FUNCTION_BLOCK T_SafeTof_Tests EXTENDS TcUnit.FB_TestSuite
VAR
    // Test_OutputDelayedOff
    group_1 : T_SafeGroup;
    fb_1 : T_SafeTof(group := group_1) := (Parameters := (DelayTime := T#100MS));
    state_1 : INT := 10;
    waitTimer_1 : TON;
    // Test_UnconnectedInputIsRefused
    group_2 : T_SafeGroup;
    fb_2 : T_SafeTof(group := group_2);
END_VAR

Test_OutputDelayedOff();
Test_UnconnectedInputIsRefused();

METHOD PRIVATE Test_OutputDelayedOff
TcUnit.TEST(__POUNAME());
waitTimer_1();

CASE state_1 OF
    10:
        group_1(Run := TRUE);
        fb_1(TofIn1 := TRUE);
        AssertEquals_BOOL(Expected := TRUE, Actual := fb_1.TofOut, Message := 'output on immediately');
        // act
        fb_1(TofIn1 := FALSE);
        AssertEquals_BOOL(Expected := TRUE, Actual := fb_1.TofOut, Message := 'output held during the delay');
        AssertEquals_BYTE(Expected := TO_BYTE(E_SafeFbState.DelayOut), Actual := fb_1.State, Message := 'state DELAYOUT');
        state_1 := 20;
        waitTimer_1(IN := TRUE, PT := T#200MS);
    20:
        group_1(Run := TRUE);
        fb_1(TofIn1 := FALSE);

        IF NOT waitTimer_1.Q THEN
            RETURN;
        END_IF

        waitTimer_1(IN := FALSE);
        // assert
        AssertEquals_BOOL(Expected := FALSE, Actual := fb_1.TofOut, Message := 'output off after the delay');
        TEST_FINISHED_NAMED(__POUNAME());
        state_1 := 10;
END_CASE
END_METHOD

METHOD PRIVATE Test_UnconnectedInputIsRefused
TcUnit.TEST(__POUNAME());
// arrange / act: TofIn1 is unconnected, which the Safety Editor refuses
group_2(Run := TRUE);
fb_2();
group_2(Run := TRUE);
fb_2();
// assert
AssertEquals_BOOL(Expected := TRUE, Actual := fb_2.Error, Message := 'configuration error reported');
AssertEquals_BYTE(Expected := TO_BYTE(E_SafeFbState.Error), Actual := fb_2.State, Message := 'state ERROR');
AssertEquals_WORD(Expected := WORD#16#8000, Actual := fb_2.Diag, Message := 'diag bit 15 configuration refused');
AssertEquals_BOOL(Expected := FALSE, Actual := fb_2.TofOut, Message := 'TofOut stays at its safe value');
AssertEquals_BOOL(Expected := TRUE, Actual := group_2.FbErr, Message := 'the group sees an FB error');
// act: ErrAck 0 -> 1 -> 0 does not clear a configuration error
group_2(Run := TRUE, ErrAck := TRUE);
fb_2();
group_2(Run := TRUE, ErrAck := TRUE);
fb_2();
group_2(Run := TRUE, ErrAck := FALSE);
fb_2();
AssertEquals_BOOL(Expected := TRUE, Actual := fb_2.Error, Message := 'error not acknowledged');
AssertEquals_WORD(Expected := WORD#16#8000, Actual := fb_2.Diag, Message := 'diag bit 15 kept');
TEST_FINISHED_NAMED(__POUNAME());
END_METHOD

END_FUNCTION_BLOCK

(* stored: Version 1.1.0.1
   POU T_SafeTof_Tests: Id {978229da-758b-5bed-80ea-cf07aeecdce2}, SpecialFunc None
   Method Test_OutputDelayedOff: Id {b6d59bd9-12c1-5814-8994-2d4710fe2757}
   Method Test_UnconnectedInputIsRefused: Id {41898d87-9230-466f-8ce4-e67e6830cca2} *)
